(* IEC 61131-3 sources: plcassist-cli/packages/volt-lsp-iec/test-corpus/pro2193/Device/Plc Logic/Application/09 Misc/Library Manager/CAA List And Tree, 21 files *)

(* ---- VERSIONCONSTANTS.gvl ---- *)
VAR_GLOBAL
	GC_BYVERSION : BYTE := 1;
	GC_BYVERSION_1 : BYTE := 0;
END_VAR

(* ---- IELEMENT.itf ---- *)
INTERFACE IELEMENT
END_INTERFACE

METHOD ISLISTMEMBEROF : BOOL
VAR_INPUT
	ITFLIST : ISimpleList;
END_VAR
END_METHOD

(* ---- IELEMENTHELPER.itf ---- *)
INTERFACE IELEMENTHELPER
END_INTERFACE

METHOD PRVREMOVEELEM : IElementHelper
END_METHOD

(* ---- ILIST.itf ---- *)
INTERFACE ILIST
END_INTERFACE

METHOD INSERTELEM : IElement
VAR_INPUT
	ITFELEMENT : IElement;
	ITFPRECURSOR : IElement;
END_VAR
END_METHOD

METHOD APPENDELEM : IElement
VAR_INPUT
	ITFELEMENT : IElement;
END_VAR
END_METHOD

METHOD REMOVEELEM : IElement
VAR_INPUT
	ITFELEMENT : IElement;
END_VAR
END_METHOD

METHOD POPELEM : IElement
END_METHOD

METHOD POPBACKELEM : IElement
END_METHOD

METHOD PUSHELEM : IElement
VAR_INPUT
	ITFELEMENT : IElement;
END_VAR
END_METHOD

(* ---- ILISTHELPER.itf ---- *)
INTERFACE ILISTHELPER
END_INTERFACE

METHOD PRVINSERTELEM : IElementHelper
VAR_INPUT
	ITFELEMENT : IElementHelper;
	ITFPRECURSOR : IElementHelper;
END_VAR
END_METHOD

METHOD PRVAPPENDELEM : IElementHelper
VAR_INPUT
	ITFELEMENT : IElementHelper;
END_VAR
END_METHOD

METHOD PRVREMOVEELEM : IElementHelper
VAR_INPUT
	ITFELEMENT : IElementHelper;
END_VAR
END_METHOD

METHOD PRVPOPELEM : IElementHelper
END_METHOD

METHOD PRVPOPBACKELEM : IElementHelper
END_METHOD

METHOD PRVPUSHELEM : IElementHelper
VAR_INPUT
	ITFELEMENT : IElementHelper;
END_VAR
END_METHOD

(* ---- ISIMPLELIST.itf ---- *)
INTERFACE ISIMPLELIST
END_INTERFACE

(* ---- ISIMPLETREE.itf ---- *)
INTERFACE ISIMPLETREE
END_INTERFACE

(* ---- ITREE.itf ---- *)
INTERFACE ITREE
END_INTERFACE

METHOD ADDCHILD : ITree
VAR_INPUT
	ITFCHILD : ITree;
	XASFIRSTCHILD : BOOL;
END_VAR
END_METHOD

METHOD INSERTSIBLING : ITree
VAR_INPUT
	ITFSIBLING : ITree;
END_VAR
END_METHOD

METHOD REMOVETREE : ITree
END_METHOD

(* ---- ITREEHELPER.itf ---- *)
INTERFACE ITREEHELPER
END_INTERFACE

METHOD PRVADDCHILD : ITreeHelper
VAR_INPUT
	ITFCHILD : ITreeHelper;
	XASFIRSTCHILD : BOOL;
END_VAR
END_METHOD

METHOD PRVINSERTSIBLING : ITreeHelper
VAR_INPUT
	ITFSIBLING : ITreeHelper;
END_VAR
END_METHOD

METHOD PRVREMOVETREE : ITreeHelper
END_METHOD

(* ---- ITYPEDELEMENT.itf ---- *)
INTERFACE ITYPEDELEMENT
END_INTERFACE

(* ---- ITYPEDLIST.itf ---- *)
INTERFACE ITYPEDLIST
END_INTERFACE

METHOD POPBACKELEM : ITypedElement
END_METHOD

METHOD PUSHELEM : ITypedElement
VAR_INPUT
	ITFELEMENT : ITypedElement;
END_VAR
END_METHOD

METHOD INSERTELEM : ITypedElement
VAR_INPUT
	ITFELEMENT : ITypedElement;
	ITFPRECURSOR : ITypedElement;
END_VAR
END_METHOD

METHOD APPENDELEM : ITypedElement
VAR_INPUT
	ITFELEMENT : ITypedElement;
END_VAR
END_METHOD

METHOD REMOVEELEM : ITypedElement
VAR_INPUT
	ITFELEMENT : ITypedElement;
END_VAR
END_METHOD

METHOD POPELEM : ITypedElement
END_METHOD

(* ---- ITYPEDTREE.itf ---- *)
INTERFACE ITYPEDTREE
END_INTERFACE

METHOD ADDCHILD : ITypedTree
VAR_INPUT
	ITFCHILD : ITypedTree;
	XASFIRSTCHILD : BOOL;
END_VAR
END_METHOD

METHOD INSERTSIBLING : ITypedTree
VAR_INPUT
	ITFSIBLING : ITypedTree;
END_VAR
END_METHOD

METHOD REMOVETREE : ITypedTree
END_METHOD

(* ---- GETSUPPLIERVERSION.fun ---- *)
FUNCTION GETSUPPLIERVERSION : WORD
END_FUNCTION

(* ---- ELEMENT.fb ---- *)
FUNCTION_BLOCK ELEMENT
VAR
	ITFPREV : IElementHelper;
	ITFNEXT : IElementHelper;
	ITFLIST : IListHelper;
	ISLINKEDELEM : BOOL;
	NEXTELEM : IElement;
	PREVELEM : IElement;
	PRVLIST : IListHelper;
	PRVNEXTELEM : IElementHelper;
	PRVPREVELEM : IElementHelper;
END_VAR
END_FUNCTION_BLOCK

METHOD ISLISTMEMBEROF : BOOL
VAR_INPUT
	ITFLIST : ISimpleList;
END_VAR
END_METHOD

METHOD PRVREMOVEELEM : IElementHelper
END_METHOD

(* ---- LIST.fb ---- *)
FUNCTION_BLOCK LIST EXTENDS ListBase
END_FUNCTION_BLOCK

METHOD APPENDELEM : IElement
VAR_INPUT
	ITFELEMENT : IElement;
END_VAR
END_METHOD

METHOD INSERTELEM : IElement
VAR_INPUT
	ITFELEMENT : IElement;
	ITFPRECURSOR : IElement;
END_VAR
END_METHOD

METHOD POPBACKELEM : IElement
END_METHOD

METHOD POPELEM : IElement
END_METHOD

METHOD PUSHELEM : IElement
VAR_INPUT
	ITFELEMENT : IElement;
END_VAR
END_METHOD

METHOD REMOVEELEM : IElement
VAR_INPUT
	ITFELEMENT : IElement;
END_VAR
END_METHOD

(* ---- LISTBASE.fb ---- *)
FUNCTION_BLOCK LISTBASE
VAR
	ITFHEAD : IElementHelper;
	ITFTAIL : IElementHelper;
	CTSIZE : CAA.COUNT;
	HEADELEM : IElement;
	LISTISEMPTY : BOOL;
	LISTSIZE : CAA.COUNT;
	TAILELEM : IElement;
END_VAR
END_FUNCTION_BLOCK

METHOD PRVAPPENDELEM : IElementHelper
VAR_INPUT
	ITFELEMENT : IElementHelper;
END_VAR
END_METHOD

METHOD PRVINSERTELEM : IElementHelper
VAR_INPUT
	ITFELEMENT : IElementHelper;
	ITFPRECURSOR : IElementHelper;
END_VAR
END_METHOD

METHOD PRVPOPBACKELEM : IElementHelper
END_METHOD

METHOD PRVPOPELEM : IElementHelper
END_METHOD

METHOD PRVPUSHELEM : IElementHelper
VAR_INPUT
	ITFELEMENT : IElementHelper;
END_VAR
END_METHOD

METHOD PRVREMOVEELEM : IElementHelper
VAR_INPUT
	ITFELEMENT : IElementHelper;
END_VAR
END_METHOD

(* ---- TREE.fb ---- *)
FUNCTION_BLOCK TREE EXTENDS TreeBase
END_FUNCTION_BLOCK

METHOD ADDCHILD : ITree
VAR_INPUT
	ITFCHILD : ITree;
	XASFIRSTCHILD : BOOL;
END_VAR
END_METHOD

METHOD INSERTSIBLING : ITree
VAR_INPUT
	ITFSIBLING : ITree;
END_VAR
END_METHOD

METHOD REMOVETREE : ITree
END_METHOD

(* ---- TREEBASE.fb ---- *)
FUNCTION_BLOCK TREEBASE
VAR
	ITFPARENT : ITreeHelper;
	ITFNEXTSIBLING : ITreeHelper;
	ITFPREVSIBLING : ITreeHelper;
	ITFFIRSTCHILD : ITreeHelper;
	ITFLASTCHILD : ITreeHelper;
	CTCHILDCOUNT : CAA.COUNT;
	CHILDCOUNT : CAA.COUNT;
	FIRSTCHILD : ISimpleTree;
	ISLINKEDTREE : BOOL;
	ISTREEROOT : BOOL;
	LASTCHILD : ISimpleTree;
	NEXTSIBLING : ISimpleTree;
	PARENTTREE : ISimpleTree;
	PREVSIBLING : ISimpleTree;
	PRVCHILDCOUNT : CAA.COUNT;
	PRVFIRSTCHILD : ITreeHelper;
	PRVLASTCHILD : ITreeHelper;
	PRVNEXTSIBLING : ITreeHelper;
	PRVPARENTTREE : ITreeHelper;
	PRVPREVSIBLING : ITreeHelper;
	SIBLINGCOUNT : CAA.COUNT;
END_VAR
END_FUNCTION_BLOCK

METHOD PRVADDCHILD : ITreeHelper
VAR_INPUT
	ITFCHILD : ITreeHelper;
	XASFIRSTCHILD : BOOL;
END_VAR
END_METHOD

METHOD PRVINSERTSIBLING : ITreeHelper
VAR_INPUT
	ITFSIBLING : ITreeHelper;
END_VAR
END_METHOD

METHOD PRVREMOVETREE : ITreeHelper
END_METHOD

(* ---- TYPEDELEMENT.fb ---- *)
FUNCTION_BLOCK TYPEDELEMENT EXTENDS Element
VAR
	IDTYPEID : CAA.IDENT;
	ELEMTYPEID : CAA.IDENT;
END_VAR
END_FUNCTION_BLOCK

(* ---- TYPEDLIST.fb ---- *)
FUNCTION_BLOCK TYPEDLIST EXTENDS ListBase
VAR
	IDTYPEID : UDINT;
	LISTTYPEID : CAA.IDENT;
END_VAR
END_FUNCTION_BLOCK

METHOD APPENDELEM : ITypedElement
VAR_INPUT
	ITFELEMENT : ITypedElement;
END_VAR
END_METHOD

METHOD INSERTELEM : ITypedElement
VAR_INPUT
	ITFELEMENT : ITypedElement;
	ITFPRECURSOR : ITypedElement;
END_VAR
END_METHOD

METHOD POPBACKELEM : ITypedElement
END_METHOD

METHOD POPELEM : ITypedElement
END_METHOD

METHOD PUSHELEM : ITypedElement
VAR_INPUT
	ITFELEMENT : ITypedElement;
END_VAR
END_METHOD

METHOD REMOVEELEM : ITypedElement
VAR_INPUT
	ITFELEMENT : ITypedElement;
END_VAR
END_METHOD

METHOD PRVCHECKELEMENT : BOOL
VAR_INPUT
	ITFELEMENT : ITypedElement;
END_VAR
END_METHOD

(* ---- TYPEDTREE.fb ---- *)
FUNCTION_BLOCK TYPEDTREE EXTENDS TreeBase
VAR
	IDTYPEID : CAA.IDENT;
	TREETYPEID : CAA.IDENT;
END_VAR
END_FUNCTION_BLOCK

METHOD ADDCHILD : ITypedTree
VAR_INPUT
	ITFCHILD : ITypedTree;
	XASFIRSTCHILD : BOOL;
END_VAR
END_METHOD

METHOD INSERTSIBLING : ITypedTree
VAR_INPUT
	ITFSIBLING : ITypedTree;
END_VAR
END_METHOD

METHOD REMOVETREE : ITypedTree
END_METHOD

METHOD PRVCHECKTREE : BOOL
VAR_INPUT
	ITFTREE : ITypedTree;
END_VAR
END_METHOD
